(* Logix 5000 project; controller CIP_14485201 vendor 1 type 14 code 216 rev 38.11; software revision 38.01; part 3 of 12 *)
(* tags used below, declared in another part *)
   Alarm_Preset_Indx : DINT;   // ALARM TIMER PRESET INDEX POSITION
   Alarm_Timer : TIMER[128];   // ALARM MSGS 1-127 DELAY TIMERS
   Alarm_Timer_Preset : DINT[128];   // ALARM TIMER PRESETS STORAGE
   Bit : BOOL[128];   // BIT
   Integer : DINT[150];   // INTEGER
   Integer_1 : ALIAS FOR Integer[1];   // RECIPE SELECTOR LIST POSITION ALIAS
   Integer_6 : ALIAS FOR Integer[6];   // EDIT RECIPES SELECTOR LIST POSITION ALIAS
   One_Shot : BOOL[128];   // ONE SHOT ARRAY
   OpCode_Pin : DINT[5];   // OPCODE PIN ARRAY
   OpCode_Word : DINT[5,97];   // OPCODE WORD ARRAY
   Panelview : INT[40];   // PANELVIEW CONTROL
   PID2_Output_Memory : REAL;   // SUPPLY FLOW PID OUTPUT MEMORY TO USE FOR BUMPLESS TRANSFER
   Process_to_CIP : Process_to_CIP;   // PROCESS SIGNALS TO CIP
   PV_Copy_Recipes_Destination : DINT;   // COPY RECIPES DESTINATION
   PV_Copy_Recipes_Duration : TIMER;   // COPY RECIPES COPY DURATION
   PV_Copy_Recipes_One_Shot : BOOL;   // COPY RECIPES REQUEST TO COPY ONE SHOT
   PV_Copy_Recipes_Request : BOOL;   // COPY RECIPES REQUEST TO COPY
   PV_Copy_Recipes_Source : DINT;
   PV_Current_Select_Step_Op : DINT;   // PANELVIEW STORES CURRENT OPCODE NUMBER OF STEP BEING EDITED FOR DISPLAY ON OPCODE LIST SCREEN
   PV_Edit_OpCode_List : DINT[24];   // PANELVIEW RECIPE EDIT OPCODE LIST
   PV_Edit_Opcode_Sel_Top_Row : DINT;   // PANELVIEW RECIPE EDIT OPCODE LIST TOP ROW #
   PV_Edit_Opcodes : DINT[300];   // PANELVIEW BUFFER TO EDIT OPCODES
   PV_Edit_Recipe_Name : STRING;   // SELECTED RECIPE TO EDIT
   PV_Edit_Recipe_Top_Row : DINT;   // PANELVIEW RECIPE EDIT TOP ROW #
   PV_Edit_Recipes : DINT[7];   // PANELVIEW RECIPE EDITING
   PV_Edit_Recipes_0 : ALIAS FOR PV_Edit_Recipes[0];   // EDIT RECIPES STEP NUMBER
   PV_Edit_Recipes_0_Prev : DINT;   // EDIT RECIPE STEP NUMBER PREVIOUS POSITION
   PV_Edit_Screen_Opcodes : DINT[25];   // PANELVIEW RECIPE EDIT DISPLAY OPCODES
   PV_Edit_Setpoints : REAL[97];   // PANELVIEW BUFFER TO EDIT SETPOINTS
   PV_Edit_Times : DINT[300];   // PANELVIEW BUFFER TO EDIT STEP TIMES
   PV_Edit_Times_Indexer : DINT;
   PV_Edit_Times_Minutes : DINT[98];
   PV_Edit_Times_Seconds : DINT[98];
   PV_Rename_Recipe_Name : STRING;   // PANELVIEW RENAME RECIPE NAME
   PV_Step_Time : DINT;   // PANELVIEW DISPLAY STEP TIME
   pv_step_time_minutes : DINT;   // PANELVIEW DISPLAY STEP TIME MINUTES
   pv_step_time_seconds : DINT;   // PANELVIEW DISPLAY STEP TIME SECONDS
   Recipe : RECIPE[41];   // RECIPES
   Recipe_Name : STRING[41];   // RECIPE NAME STORAGE
   Recipe_Name_Indx : DINT;   // RECIPE NAME INDEX POSITION
   Recipe_Step_Length : CONTROL;   // CURRENT RECIPE LENGTH
   Sequencer : CONTROL[4];   // SEQUENCER
   Step_Time_Preset : DINT;
   Subsequent_OpCode_Pin : DINT[5];   // OPCODE PIN ARRAY
   TemporaryRecipeSelection : DINT;
   Time_Date : DINT[20];   // SYSTEM TIME/DATE EDIT/STORAGE
   Timer : TIMER[99];   // TIMER
   Timer_Chem1_Pump : TIMER[7];   // CHEM #1 CONTROL TIMERS
   Timer_Chem2_Pump : TIMER[7];   // CHEM #2 CONTROL TIMERS
   User_Security_Name_Display : STRING;

PROGRAM MainProgram   (* main routine _02_SUB *)

ROUTINE _02_SUB   (* ladder *)
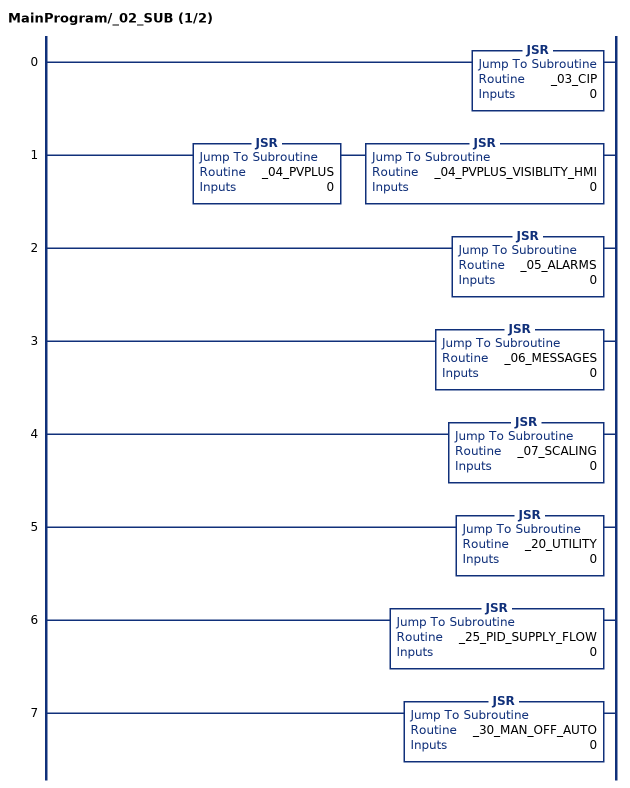
   0: JSR(_03_CIP,0);
   1: JSR(_04_PVPLUS,0)JSR(_04_PVPLUS_VISIBLITY_HMI,0);
   2: JSR(_05_ALARMS,0);
   3: JSR(_06_MESSAGES,0);
   4: JSR(_07_SCALING,0);
   5: JSR(_20_UTILITY,0);
   6: JSR(_25_PID_SUPPLY_FLOW,0);
   7: JSR(_30_MAN_OFF_AUTO,0);
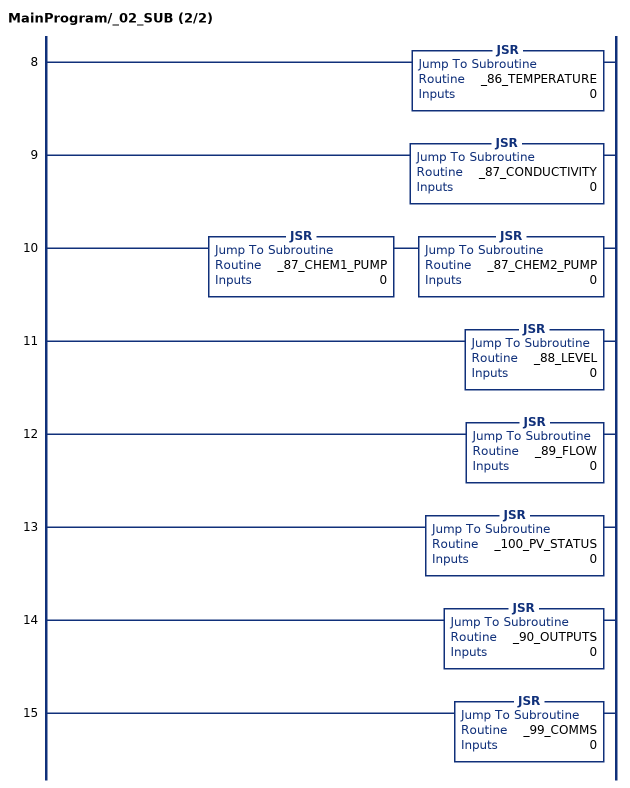
   8: JSR(_86_TEMPERATURE,0);
   9: JSR(_87_CONDUCTIVITY,0);
   10: JSR(_87_CHEM1_PUMP,0)JSR(_87_CHEM2_PUMP,0);
   11: JSR(_88_LEVEL,0);
   12: JSR(_89_FLOW,0);
   13: JSR(_100_PV_STATUS,0);
   14: JSR(_90_OUTPUTS,0);
   15: JSR(_99_COMMS,0);
END_ROUTINE

ROUTINE _03_CIP   (* ladder *)
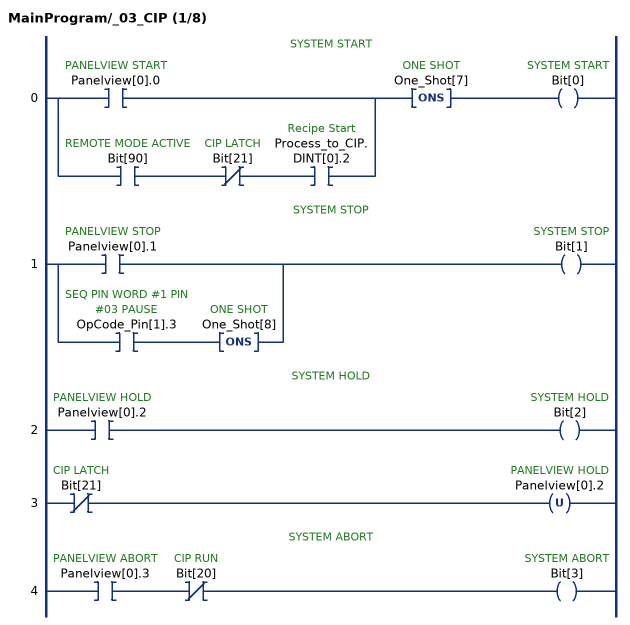
   // SYSTEM START
   0: [XIC(Panelview[0].0) ,XIC(Bit[90]) XIO(Bit[21]) XIC(Process_to_CIP.DINT[0].2) ]ONS(One_Shot[7])OTE(Bit[0]);
   // SYSTEM STOP
   1: [XIC(Panelview[0].1) ,XIC(OpCode_Pin[1].3) ONS(One_Shot[8]) ]OTE(Bit[1]);
   // SYSTEM HOLD
   2: XIC(Panelview[0].2)OTE(Bit[2]);
   3: XIO(Bit[21])OTU(Panelview[0].2);
   // SYSTEM ABORT
   4: XIC(Panelview[0].3)XIO(Bit[20])OTE(Bit[3]);
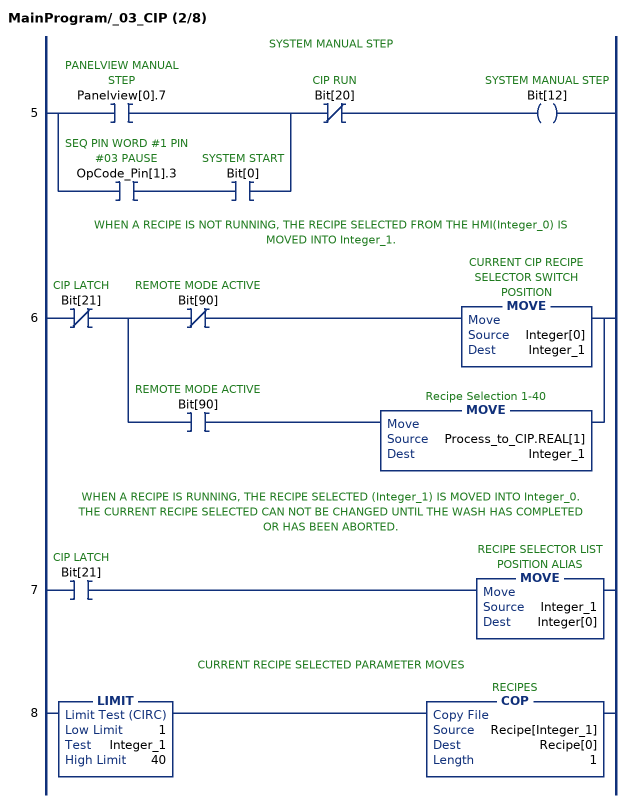
   // SYSTEM MANUAL STEP
   5: [XIC(Panelview[0].7) ,XIC(OpCode_Pin[1].3) XIC(Bit[0]) ]XIO(Bit[20])OTE(Bit[12]);
   // WHEN A RECIPE IS NOT RUNNING, THE RECIPE SELECTED FROM THE HMI(Integer_0) IS MOVED INTO Integer_1.
   6: XIO(Bit[21])[XIO(Bit[90]) MOVE(Integer[0],Integer_1) ,XIC(Bit[90]) MOVE(Process_to_CIP.REAL[1],Integer_1) ];
   // WHEN A RECIPE IS RUNNING, THE RECIPE SELECTED (Integer_1) IS MOVED INTO Integer_0.
   // THE CURRENT RECIPE SELECTED CAN NOT BE CHANGED UNTIL THE WASH HAS COMPLETED OR HAS BEEN ABORTED.
   7: XIC(Bit[21])MOVE(Integer_1,Integer[0]);
   // CURRENT RECIPE SELECTED PARAMETER MOVES
   8: LIMIT(1,Integer_1,40)COP(Recipe[Integer_1],Recipe[0],1);
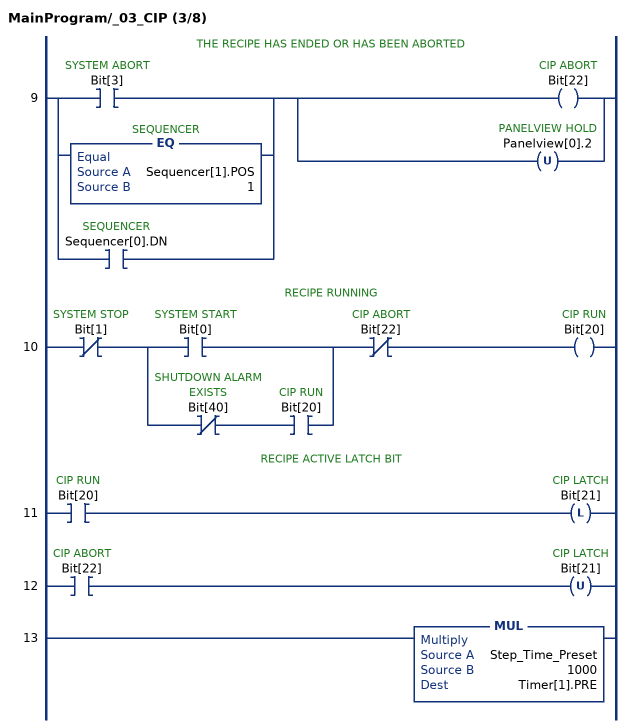
   // THE RECIPE HAS ENDED OR HAS BEEN ABORTED
   9: [XIC(Bit[3]) ,EQ(Sequencer[1].POS,1) ,XIC(Sequencer[0].DN) ][OTE(Bit[22]) ,OTU(Panelview[0].2) ];
   // RECIPE RUNNING
   10: XIO(Bit[1])[XIC(Bit[0]) ,XIO(Bit[40]) XIC(Bit[20]) ]XIO(Bit[22])OTE(Bit[20]);
   // RECIPE ACTIVE LATCH BIT
   11: XIC(Bit[20])OTL(Bit[21]);
   12: XIC(Bit[22])OTU(Bit[21]);
   13: MUL(Step_Time_Preset,1000,Timer[1].PRE);
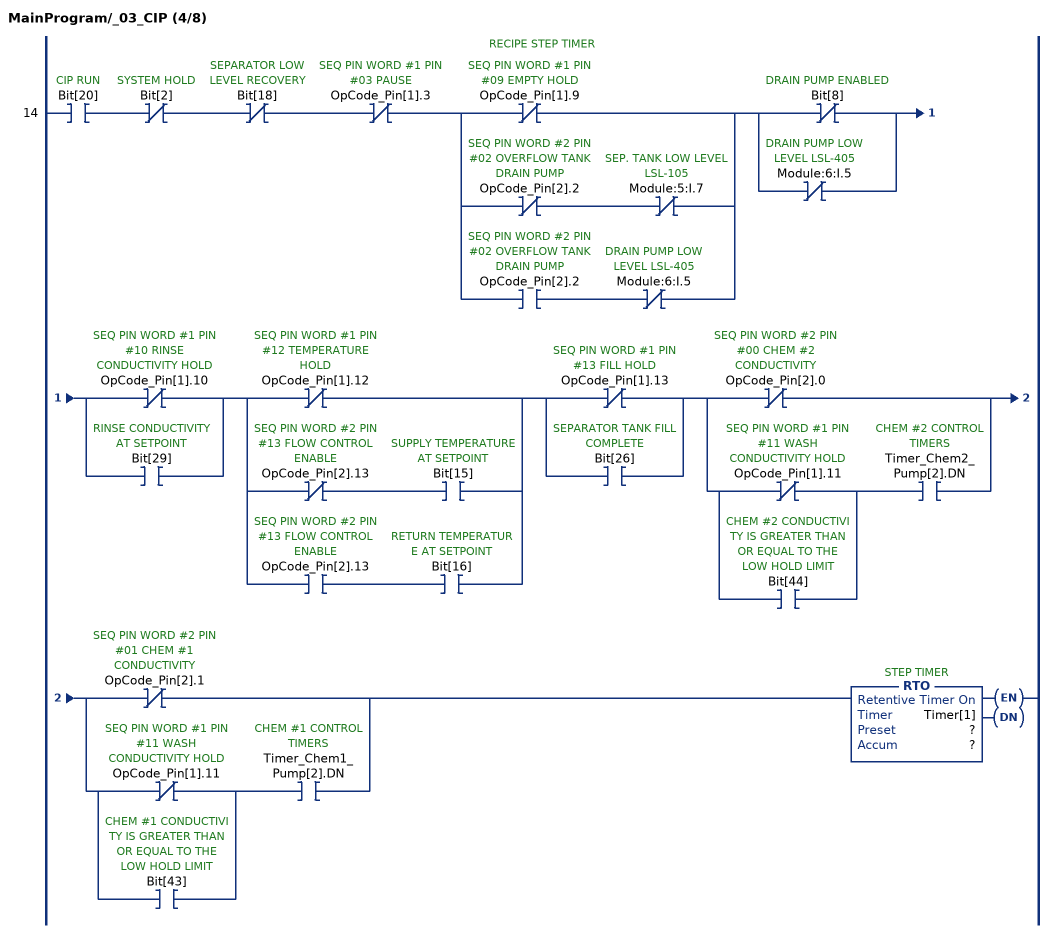
   // RECIPE STEP TIMER
   14: XIC(Bit[20])XIO(Bit[2])XIO(Bit[18])XIO(OpCode_Pin[1].3)[XIO(OpCode_Pin[1].9) ,XIO(OpCode_Pin[2].2) XIO(Module:5:I.7) ,XIC(OpCode_Pin[2].2) XIO(Module:6:I.5) ][XIO(Bit[8]) ,XIO(Module:6:I.5) ][XIO(OpCode_Pin[1].10) ,XIC(Bit[29]) ][XIO(OpCode_Pin[1].12) ,XIO(OpCode_Pin[2].13) XIC(Bit[15]) ,XIC(OpCode_Pin[2].13) XIC(Bit[16]) ][XIO(OpCode_Pin[1].13) ,XIC(Bit[26]) ][XIO(OpCode_Pin[2].0) ,[XIO(OpCode_Pin[1].11) ,XIC(Bit[44]) ] XIC(Timer_Chem2_Pump[2].DN) ][XIO(OpCode_Pin[2].1) ,[XIO(OpCode_Pin[1].11) ,XIC(Bit[43]) ] XIC(Timer_Chem1_Pump[2].DN) ]RTO(Timer[1],?,?);
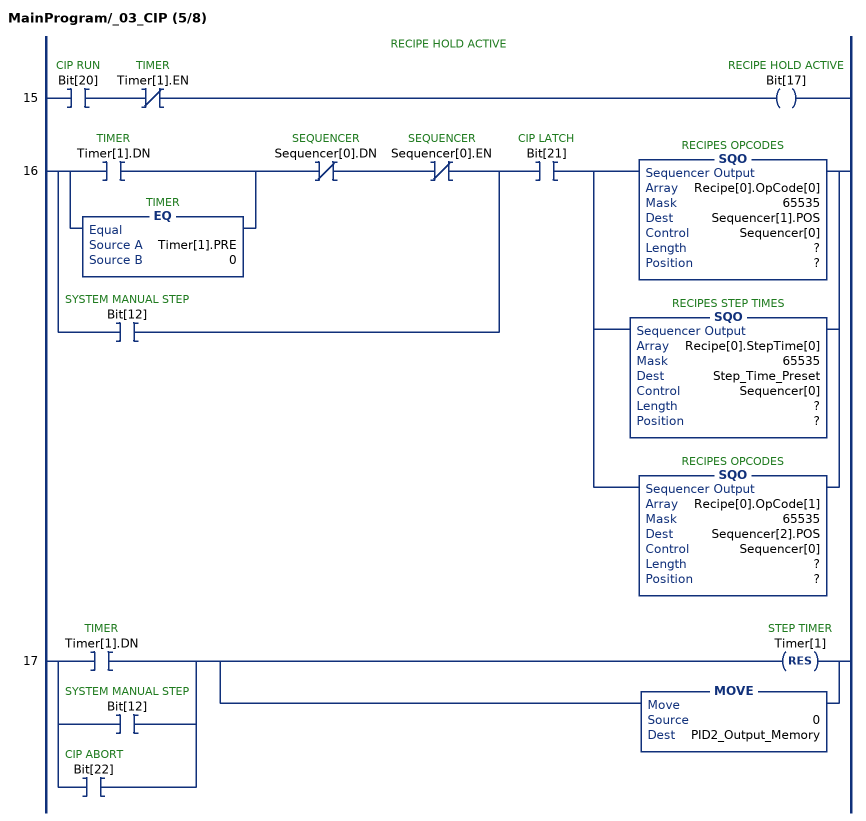
   // RECIPE HOLD ACTIVE
   15: XIC(Bit[20])XIO(Timer[1].EN)OTE(Bit[17]);
   16: [[XIC(Timer[1].DN) ,EQ(Timer[1].PRE,0) ] XIO(Sequencer[0].DN) XIO(Sequencer[0].EN) ,XIC(Bit[12]) ]XIC(Bit[21])[SQO(Recipe[0].OpCode[0],65535,Sequencer[1].POS,Sequencer[0],?,?) ,SQO(Recipe[0].StepTime[0],65535,Step_Time_Preset,Sequencer[0],?,?) ,SQO(Recipe[0].OpCode[1],65535,Sequencer[2].POS,Sequencer[0],?,?) ];
   17: [XIC(Timer[1].DN) ,XIC(Bit[12]) ,XIC(Bit[22]) ][RES(Timer[1]) ,MOVE(0,PID2_Output_Memory) ];
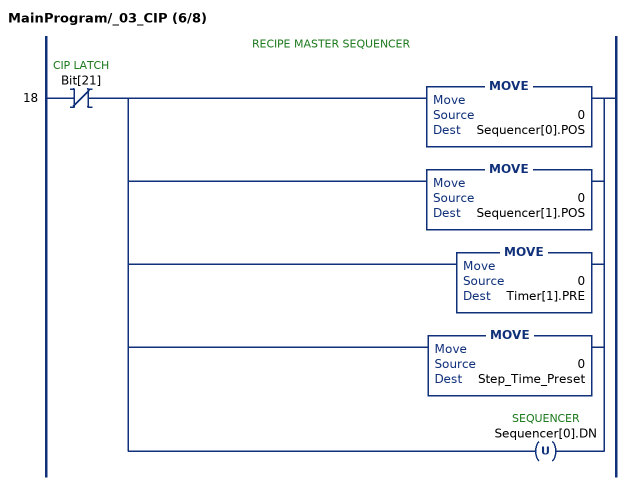
   // RECIPE MASTER SEQUENCER
   18: XIO(Bit[21])[MOVE(0,Sequencer[0].POS) ,MOVE(0,Sequencer[1].POS) ,MOVE(0,Timer[1].PRE) ,MOVE(0,Step_Time_Preset) ,OTU(Sequencer[0].DN) ];
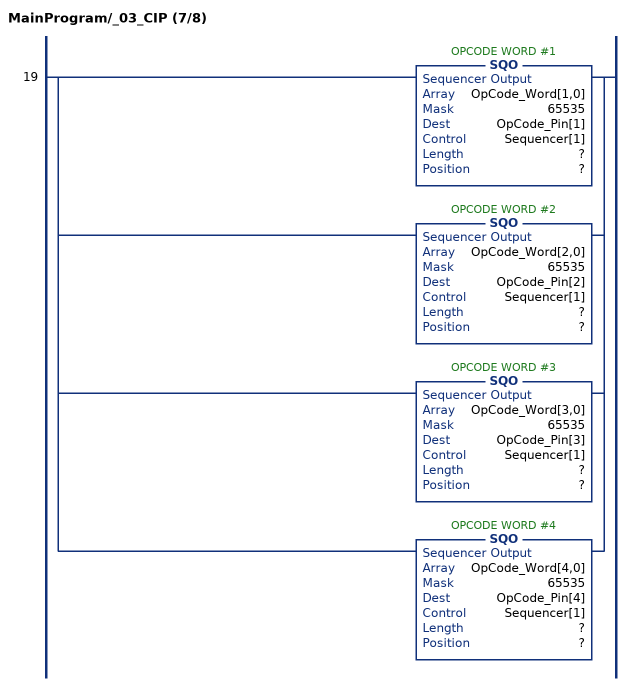
   19: [SQO(OpCode_Word[1,0],65535,OpCode_Pin[1],Sequencer[1],?,?) ,SQO(OpCode_Word[2,0],65535,OpCode_Pin[2],Sequencer[1],?,?) ,SQO(OpCode_Word[3,0],65535,OpCode_Pin[3],Sequencer[1],?,?) ,SQO(OpCode_Word[4,0],65535,OpCode_Pin[4],Sequencer[1],?,?) ];
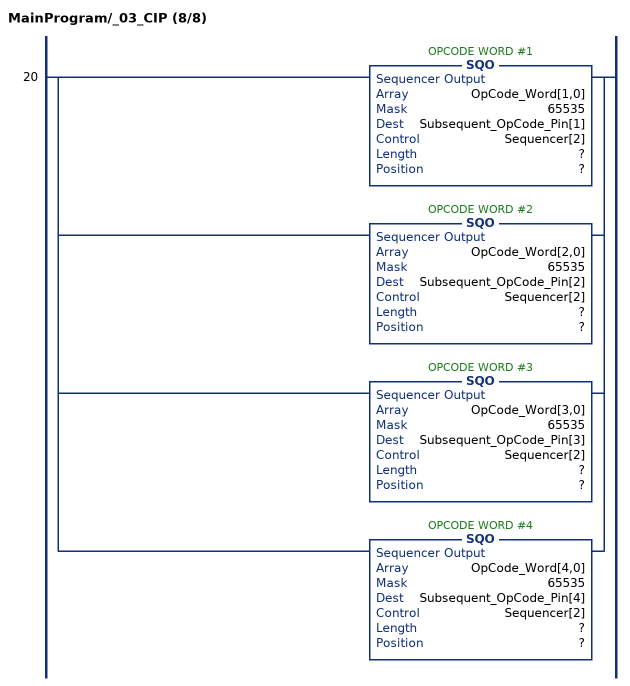
   20: [SQO(OpCode_Word[1,0],65535,Subsequent_OpCode_Pin[1],Sequencer[2],?,?) ,SQO(OpCode_Word[2,0],65535,Subsequent_OpCode_Pin[2],Sequencer[2],?,?) ,SQO(OpCode_Word[3,0],65535,Subsequent_OpCode_Pin[3],Sequencer[2],?,?) ,SQO(OpCode_Word[4,0],65535,Subsequent_OpCode_Pin[4],Sequencer[2],?,?) ];
END_ROUTINE

ROUTINE _04_PVPLUS   (* ladder *)
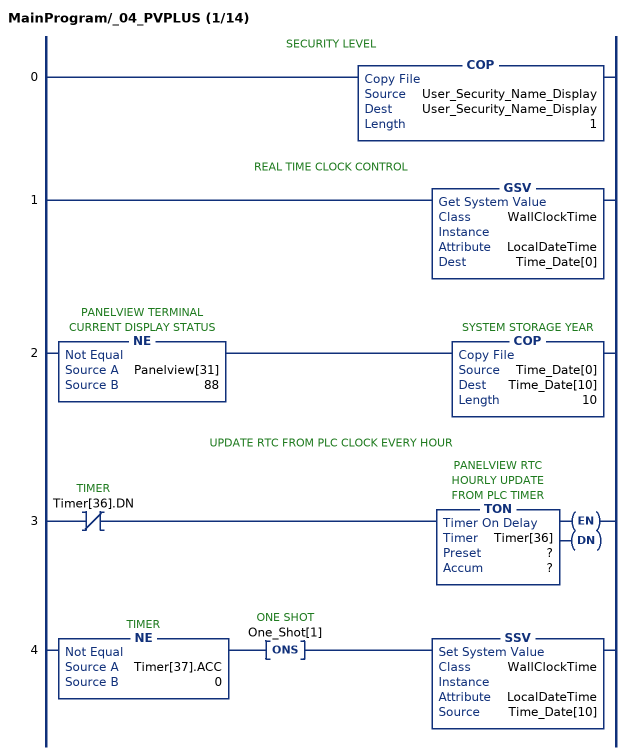
   // SECURITY LEVEL
   0: COP(User_Security_Name_Display,User_Security_Name_Display,1);
   // REAL TIME CLOCK CONTROL
   1: GSV(WallClockTime,,LocalDateTime,Time_Date[0]);
   2: NE(Panelview[31],88)COP(Time_Date[0],Time_Date[10],10);
   // UPDATE RTC FROM PLC CLOCK EVERY HOUR
   3: XIO(Timer[36].DN)TON(Timer[36],?,?);
   4: NE(Timer[37].ACC,0)ONS(One_Shot[1])SSV(WallClockTime,,LocalDateTime,Time_Date[10]);
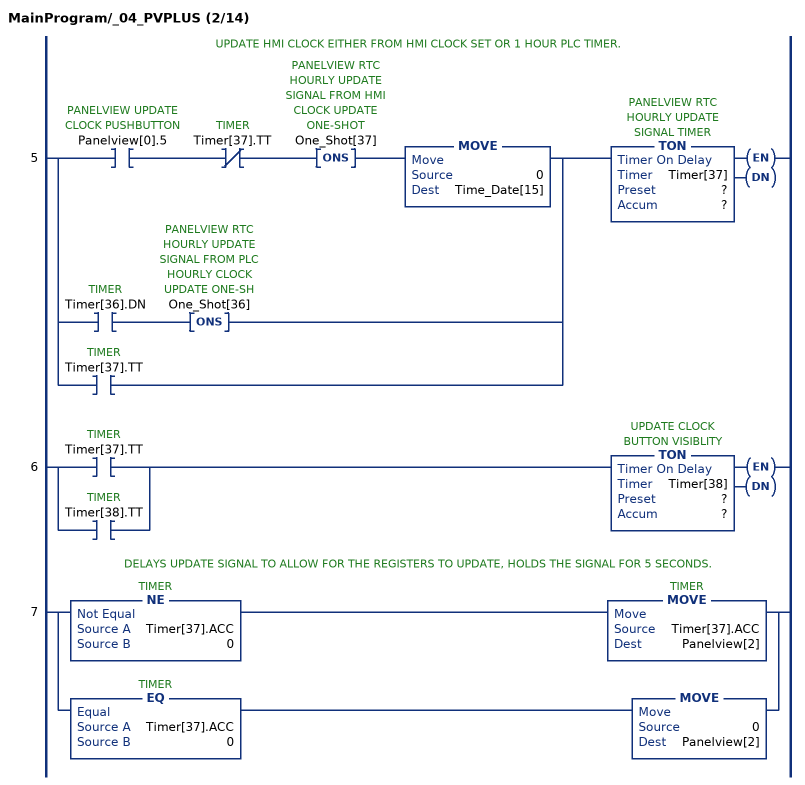
   // UPDATE HMI CLOCK EITHER FROM HMI CLOCK SET OR 1 HOUR PLC TIMER.
   5: [XIC(Panelview[0].5) XIO(Timer[37].TT) ONS(One_Shot[37]) MOVE(0,Time_Date[15]) ,XIC(Timer[36].DN) ONS(One_Shot[36]) ,XIC(Timer[37].TT) ]TON(Timer[37],?,?);
   6: [XIC(Timer[37].TT) ,XIC(Timer[38].TT) ]TON(Timer[38],?,?);
   // DELAYS UPDATE SIGNAL TO ALLOW FOR THE REGISTERS TO UPDATE, HOLDS THE SIGNAL FOR 5 SECONDS.
   7: [NE(Timer[37].ACC,0) MOVE(Timer[37].ACC,Panelview[2]) ,EQ(Timer[37].ACC,0) MOVE(0,Panelview[2]) ];
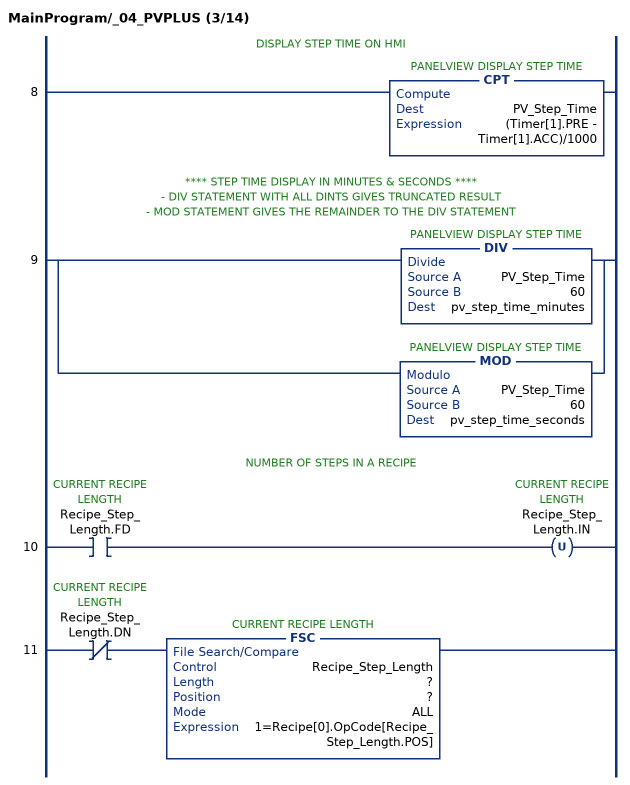
   // DISPLAY STEP TIME ON HMI
   8: CPT(PV_Step_Time,(Timer[1].PRE - Timer[1].ACC)/1000);
   // **** STEP TIME DISPLAY IN MINUTES & SECONDS ****
   // - DIV STATEMENT WITH ALL DINTS GIVES TRUNCATED RESULT
   // - MOD STATEMENT GIVES THE REMAINDER TO THE DIV STATEMENT
   9: [DIV(PV_Step_Time,60,pv_step_time_minutes) ,MOD(PV_Step_Time,60,pv_step_time_seconds) ];
   // NUMBER OF STEPS IN A RECIPE
   10: XIC(Recipe_Step_Length.FD)OTU(Recipe_Step_Length.IN);
   11: XIO(Recipe_Step_Length.DN)FSC(Recipe_Step_Length,?,?,ALL,1=Recipe[0].OpCode[Recipe_Step_Length.POS]);
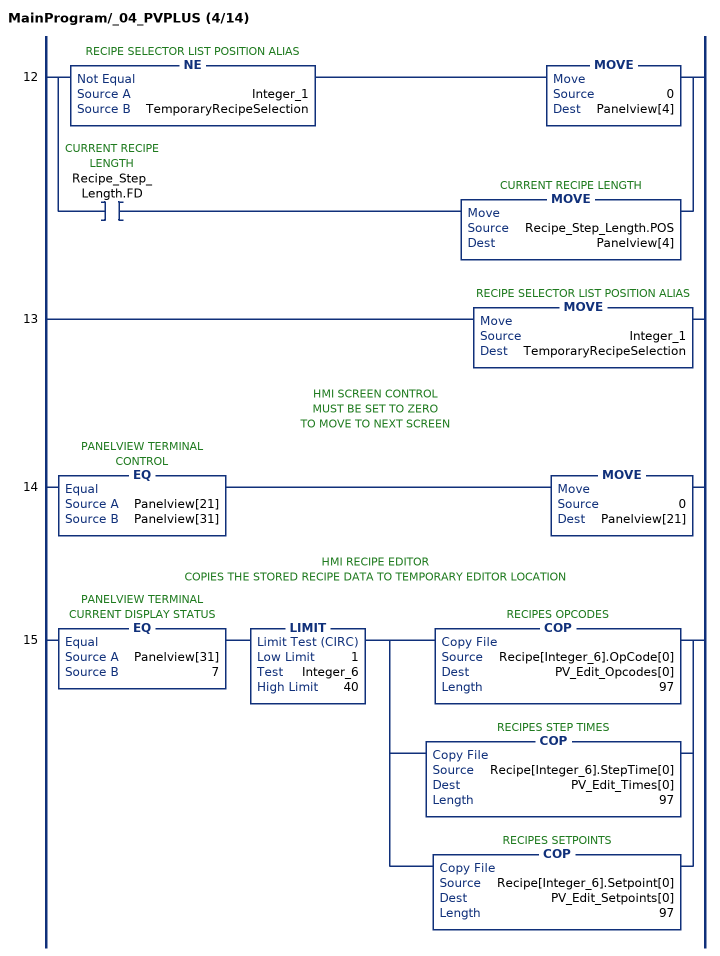
   12: [NE(Integer_1,TemporaryRecipeSelection) MOVE(0,Panelview[4]) ,XIC(Recipe_Step_Length.FD) MOVE(Recipe_Step_Length.POS,Panelview[4]) ];
   13: MOVE(Integer_1,TemporaryRecipeSelection);
   // HMI SCREEN CONTROL
   // MUST BE SET TO ZERO
   // TO MOVE TO NEXT SCREEN
   14: EQ(Panelview[21],Panelview[31])MOVE(0,Panelview[21]);
   // HMI RECIPE EDITOR
   // COPIES THE STORED RECIPE DATA TO TEMPORARY EDITOR LOCATION
   15: EQ(Panelview[31],7)LIMIT(1,Integer_6,40)[COP(Recipe[Integer_6].OpCode[0],PV_Edit_Opcodes[0],97) ,COP(Recipe[Integer_6].StepTime[0],PV_Edit_Times[0],97) ,COP(Recipe[Integer_6].Setpoint[0],PV_Edit_Setpoints[0],97) ];
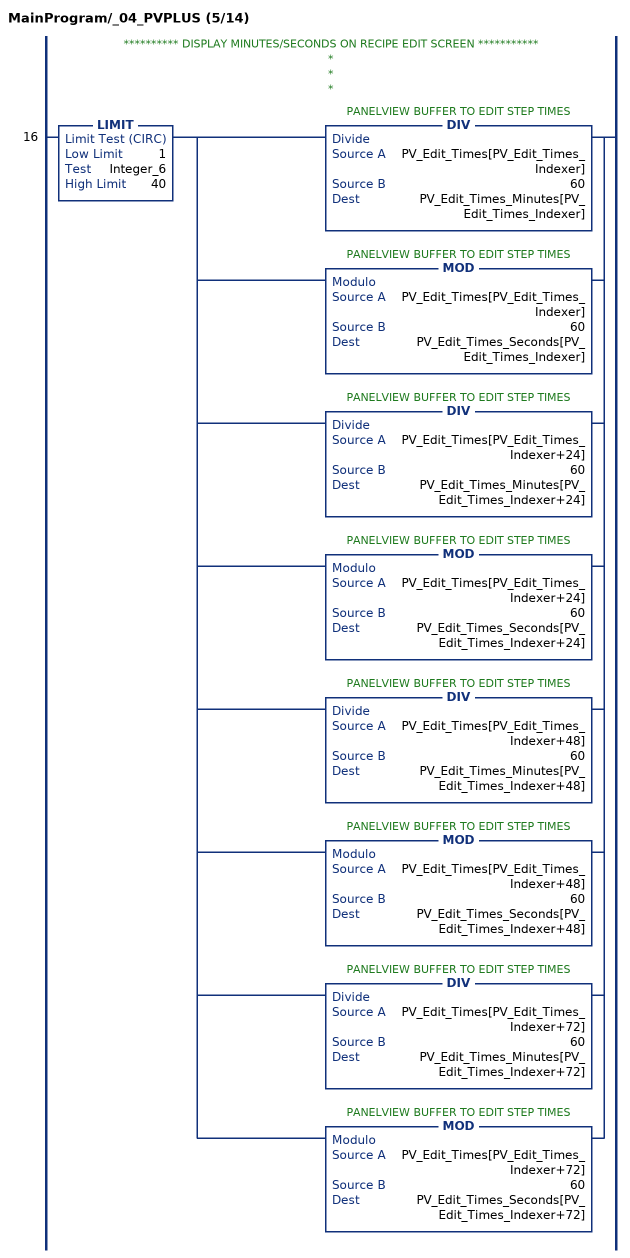
   // ********** DISPLAY MINUTES/SECONDS ON RECIPE EDIT SCREEN ***********
   // *
   // *
   // *
   16: LIMIT(1,Integer_6,40)[DIV(PV_Edit_Times[PV_Edit_Times_Indexer],60,PV_Edit_Times_Minutes[PV_Edit_Times_Indexer]) ,MOD(PV_Edit_Times[PV_Edit_Times_Indexer],60,PV_Edit_Times_Seconds[PV_Edit_Times_Indexer]) ,DIV(PV_Edit_Times[PV_Edit_Times_Indexer+24],60,PV_Edit_Times_Minutes[PV_Edit_Times_Indexer+24]) ,MOD(PV_Edit_Times[PV_Edit_Times_Indexer+24],60,PV_Edit_Times_Seconds[PV_Edit_Times_Indexer+24]) ,DIV(PV_Edit_Times[PV_Edit_Times_Indexer+48],60,PV_Edit_Times_Minutes[PV_Edit_Times_Indexer+48]) ,MOD(PV_Edit_Times[PV_Edit_Times_Indexer+48],60,PV_Edit_Times_Seconds[PV_Edit_Times_Indexer+48]) ,DIV(PV_Edit_Times[PV_Edit_Times_Indexer+72],60,PV_Edit_Times_Minutes[PV_Edit_Times_Indexer+72]) ,MOD(PV_Edit_Times[PV_Edit_Times_Indexer+72],60,PV_Edit_Times_Seconds[PV_Edit_Times_Indexer+72]) ];
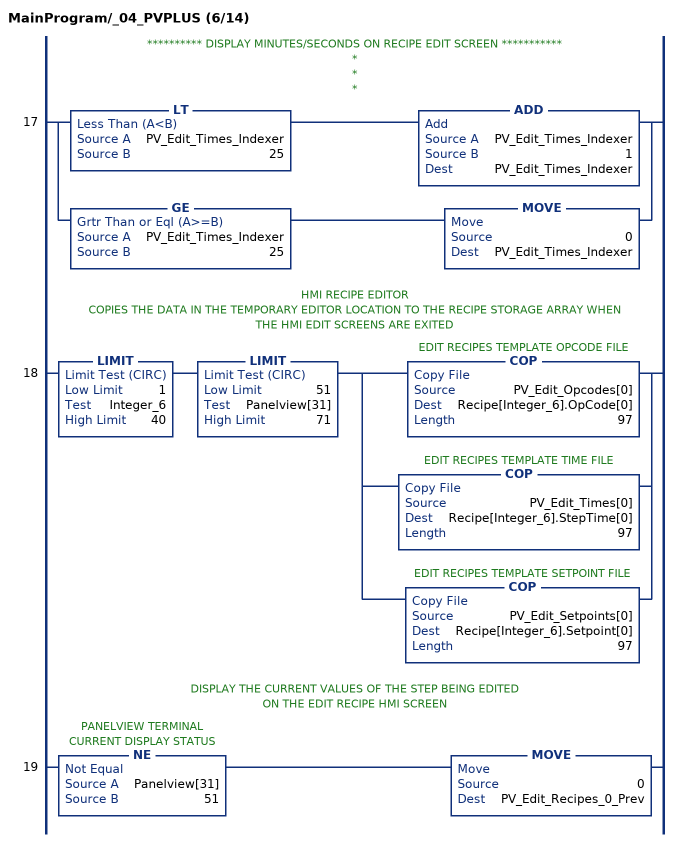
   // ********** DISPLAY MINUTES/SECONDS ON RECIPE EDIT SCREEN ***********
   // *
   // *
   // *
   17: [LT(PV_Edit_Times_Indexer,25) ADD(PV_Edit_Times_Indexer,1,PV_Edit_Times_Indexer) ,GE(PV_Edit_Times_Indexer,25) MOVE(0,PV_Edit_Times_Indexer) ];
   // HMI RECIPE EDITOR
   // COPIES THE DATA IN THE TEMPORARY EDITOR LOCATION TO THE RECIPE STORAGE ARRAY WHEN THE HMI EDIT SCREENS ARE EXITED
   18: LIMIT(1,Integer_6,40)LIMIT(51,Panelview[31],71)[COP(PV_Edit_Opcodes[0],Recipe[Integer_6].OpCode[0],97) ,COP(PV_Edit_Times[0],Recipe[Integer_6].StepTime[0],97) ,COP(PV_Edit_Setpoints[0],Recipe[Integer_6].Setpoint[0],97) ];
   // DISPLAY THE CURRENT VALUES OF THE STEP BEING EDITED
   // ON THE EDIT RECIPE HMI SCREEN
   19: NE(Panelview[31],51)MOVE(0,PV_Edit_Recipes_0_Prev);
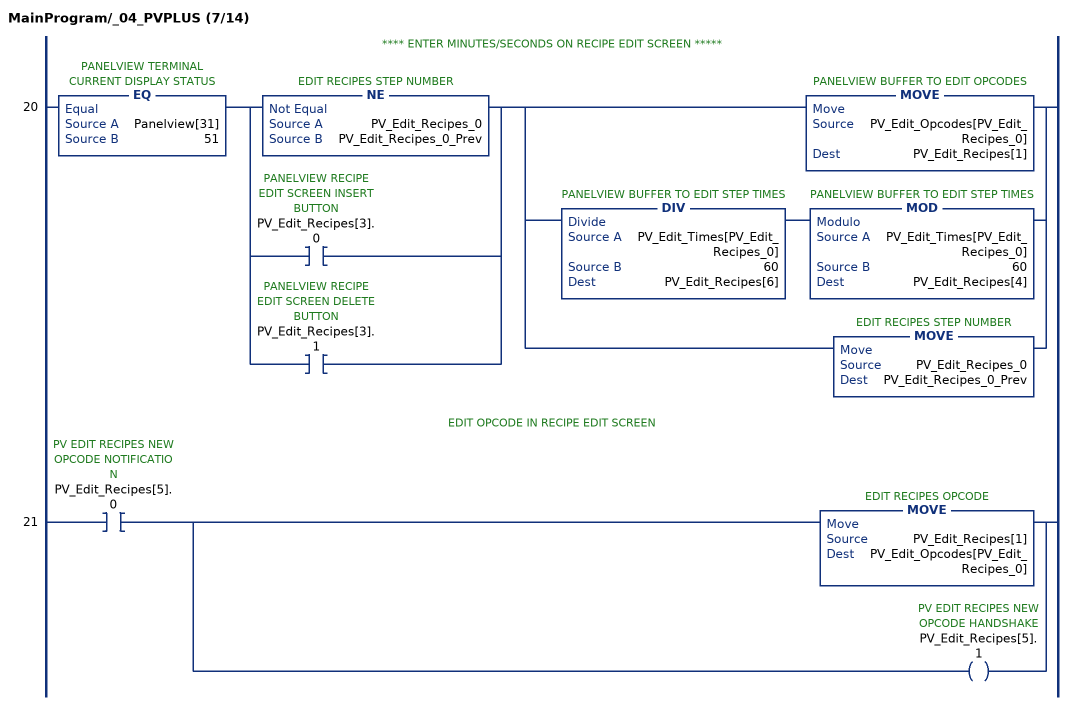
   // **** ENTER MINUTES/SECONDS ON RECIPE EDIT SCREEN *****
   20: EQ(Panelview[31],51)[NE(PV_Edit_Recipes_0,PV_Edit_Recipes_0_Prev) ,XIC(PV_Edit_Recipes[3].0) ,XIC(PV_Edit_Recipes[3].1) ][MOVE(PV_Edit_Opcodes[PV_Edit_Recipes_0],PV_Edit_Recipes[1]) ,DIV(PV_Edit_Times[PV_Edit_Recipes_0],60,PV_Edit_Recipes[6]) MOD(PV_Edit_Times[PV_Edit_Recipes_0],60,PV_Edit_Recipes[4]) ,MOVE(PV_Edit_Recipes_0,PV_Edit_Recipes_0_Prev) ];
   // EDIT OPCODE IN RECIPE EDIT SCREEN
   21: XIC(PV_Edit_Recipes[5].0)[MOVE(PV_Edit_Recipes[1],PV_Edit_Opcodes[PV_Edit_Recipes_0]) ,OTE(PV_Edit_Recipes[5].1) ];
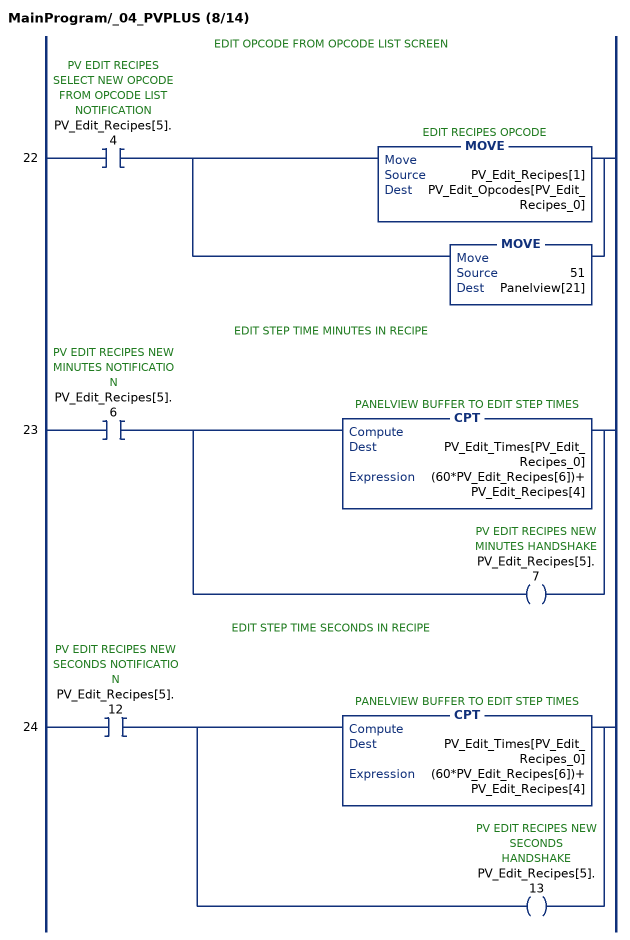
   // EDIT OPCODE FROM OPCODE LIST SCREEN
   22: XIC(PV_Edit_Recipes[5].4)[MOVE(PV_Edit_Recipes[1],PV_Edit_Opcodes[PV_Edit_Recipes_0]) ,MOVE(51,Panelview[21]) ];
   // EDIT STEP TIME MINUTES IN RECIPE
   23: XIC(PV_Edit_Recipes[5].6)[CPT(PV_Edit_Times[PV_Edit_Recipes_0],(60*PV_Edit_Recipes[6])+ PV_Edit_Recipes[4]) ,OTE(PV_Edit_Recipes[5].7) ];
   // EDIT STEP TIME SECONDS IN RECIPE
   24: XIC(PV_Edit_Recipes[5].12)[CPT(PV_Edit_Times[PV_Edit_Recipes_0],(60*PV_Edit_Recipes[6])+ PV_Edit_Recipes[4]) ,OTE(PV_Edit_Recipes[5].13) ];
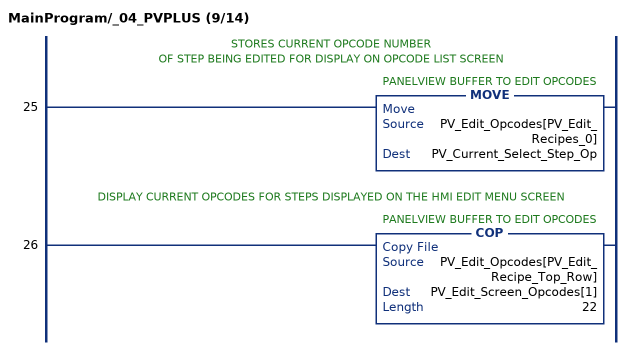
   // STORES CURRENT OPCODE NUMBER
   // OF STEP BEING EDITED FOR DISPLAY ON OPCODE LIST SCREEN
   25: MOVE(PV_Edit_Opcodes[PV_Edit_Recipes_0],PV_Current_Select_Step_Op);
   // DISPLAY CURRENT OPCODES FOR STEPS DISPLAYED ON THE HMI EDIT MENU SCREEN
   26: COP(PV_Edit_Opcodes[PV_Edit_Recipe_Top_Row],PV_Edit_Screen_Opcodes[1],22);
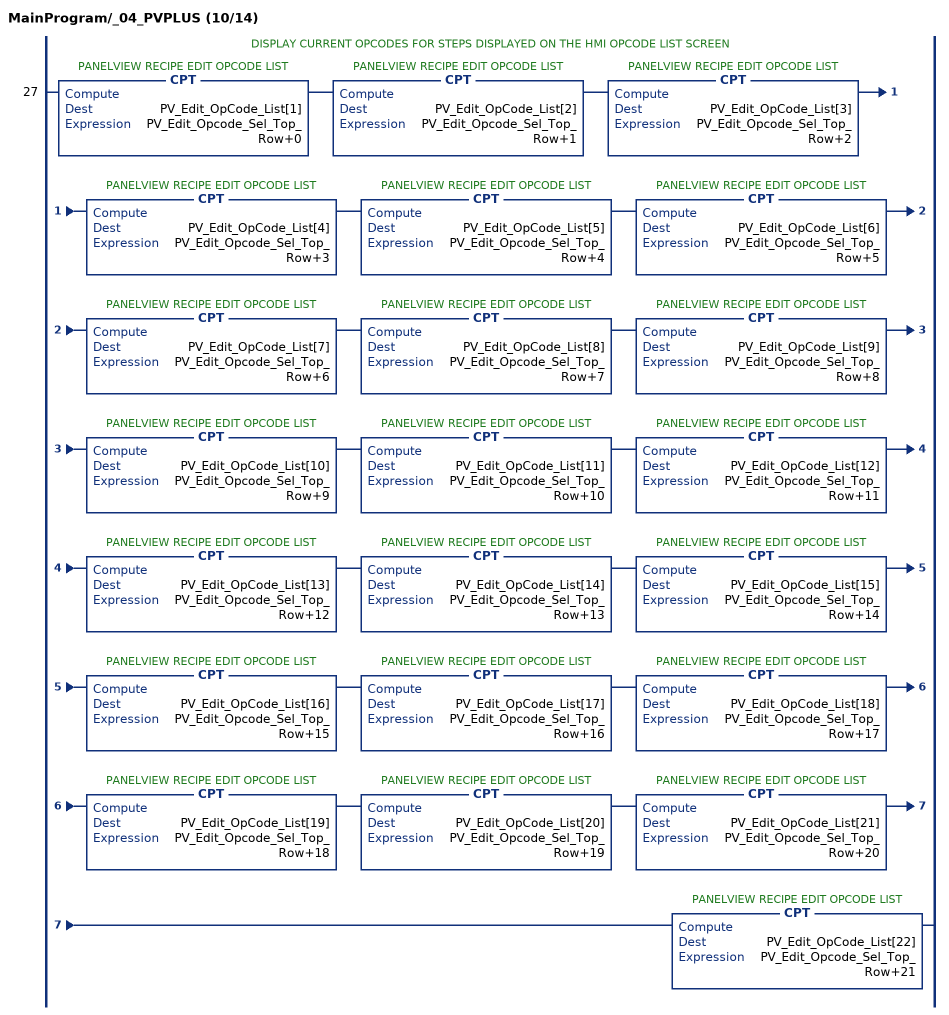
   // DISPLAY CURRENT OPCODES FOR STEPS DISPLAYED ON THE HMI OPCODE LIST SCREEN
   27: CPT(PV_Edit_OpCode_List[1],PV_Edit_Opcode_Sel_Top_Row+0)CPT(PV_Edit_OpCode_List[2],PV_Edit_Opcode_Sel_Top_Row+1)CPT(PV_Edit_OpCode_List[3],PV_Edit_Opcode_Sel_Top_Row+2)CPT(PV_Edit_OpCode_List[4],PV_Edit_Opcode_Sel_Top_Row+3)CPT(PV_Edit_OpCode_List[5],PV_Edit_Opcode_Sel_Top_Row+4)CPT(PV_Edit_OpCode_List[6],PV_Edit_Opcode_Sel_Top_Row+5)CPT(PV_Edit_OpCode_List[7],PV_Edit_Opcode_Sel_Top_Row+6)CPT(PV_Edit_OpCode_List[8],PV_Edit_Opcode_Sel_Top_Row+7)CPT(PV_Edit_OpCode_List[9],PV_Edit_Opcode_Sel_Top_Row+8)CPT(PV_Edit_OpCode_List[10],PV_Edit_Opcode_Sel_Top_Row+9)CPT(PV_Edit_OpCode_List[11],PV_Edit_Opcode_Sel_Top_Row+10)CPT(PV_Edit_OpCode_List[12],PV_Edit_Opcode_Sel_Top_Row+11)CPT(PV_Edit_OpCode_List[13],PV_Edit_Opcode_Sel_Top_Row+12)CPT(PV_Edit_OpCode_List[14],PV_Edit_Opcode_Sel_Top_Row+13)CPT(PV_Edit_OpCode_List[15],PV_Edit_Opcode_Sel_Top_Row+14)CPT(PV_Edit_OpCode_List[16],PV_Edit_Opcode_Sel_Top_Row+15)CPT(PV_Edit_OpCode_List[17],PV_Edit_Opcode_Sel_Top_Row+16)CPT(PV_Edit_OpCode_List[18],PV_Edit_Opcode_Sel_Top_Row+17)CPT(PV_Edit_OpCode_List[19],PV_Edit_Opcode_Sel_Top_Row+18)CPT(PV_Edit_OpCode_List[20],PV_Edit_Opcode_Sel_Top_Row+19)CPT(PV_Edit_OpCode_List[21],PV_Edit_Opcode_Sel_Top_Row+20)CPT(PV_Edit_OpCode_List[22],PV_Edit_Opcode_Sel_Top_Row+21);
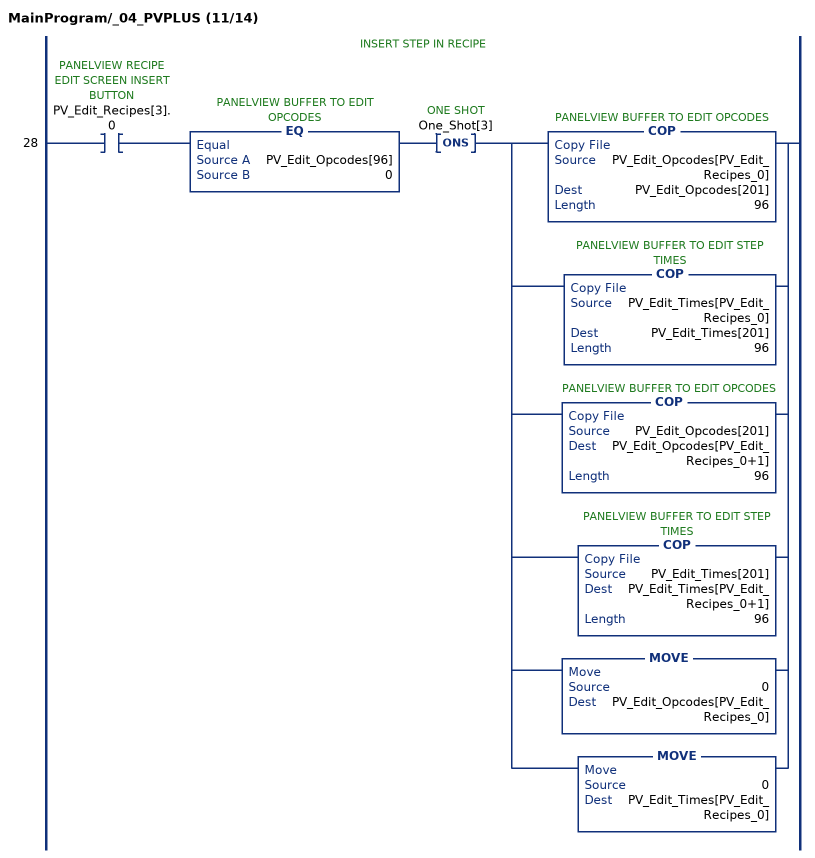
   // INSERT STEP IN RECIPE
   28: XIC(PV_Edit_Recipes[3].0)EQ(PV_Edit_Opcodes[96],0)ONS(One_Shot[3])[COP(PV_Edit_Opcodes[PV_Edit_Recipes_0],PV_Edit_Opcodes[201],96) ,COP(PV_Edit_Times[PV_Edit_Recipes_0],PV_Edit_Times[201],96) ,COP(PV_Edit_Opcodes[201],PV_Edit_Opcodes[PV_Edit_Recipes_0+1],96) ,COP(PV_Edit_Times[201],PV_Edit_Times[PV_Edit_Recipes_0+1],96) ,MOVE(0,PV_Edit_Opcodes[PV_Edit_Recipes_0]) ,MOVE(0,PV_Edit_Times[PV_Edit_Recipes_0]) ];
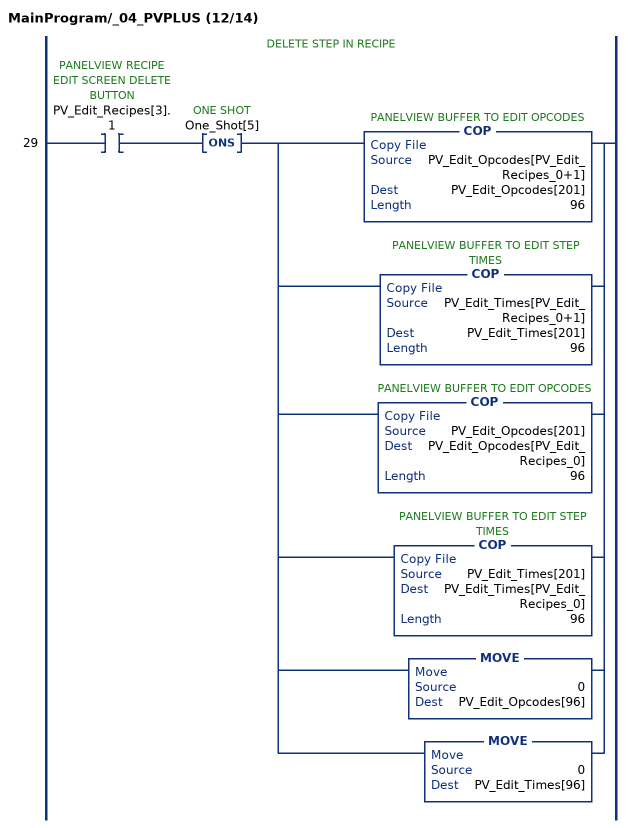
   // DELETE STEP IN RECIPE
   29: XIC(PV_Edit_Recipes[3].1)ONS(One_Shot[5])[COP(PV_Edit_Opcodes[PV_Edit_Recipes_0+1],PV_Edit_Opcodes[201],96) ,COP(PV_Edit_Times[PV_Edit_Recipes_0+1],PV_Edit_Times[201],96) ,COP(PV_Edit_Opcodes[201],PV_Edit_Opcodes[PV_Edit_Recipes_0],96) ,COP(PV_Edit_Times[201],PV_Edit_Times[PV_Edit_Recipes_0],96) ,MOVE(0,PV_Edit_Opcodes[96]) ,MOVE(0,PV_Edit_Times[96]) ];
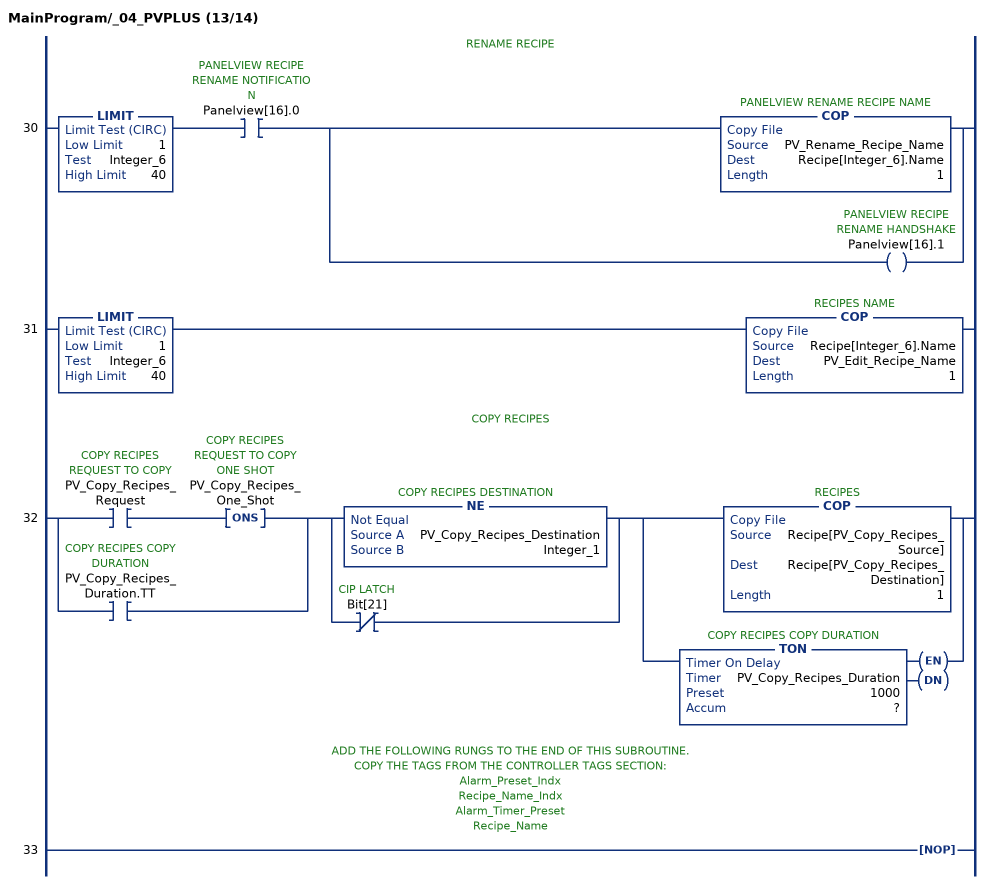
   // RENAME RECIPE
   30: LIMIT(1,Integer_6,40)XIC(Panelview[16].0)[COP(PV_Rename_Recipe_Name,Recipe[Integer_6].Name,1) ,OTE(Panelview[16].1) ];
   31: LIMIT(1,Integer_6,40)COP(Recipe[Integer_6].Name,PV_Edit_Recipe_Name,1);
   // COPY RECIPES
   32: [XIC(PV_Copy_Recipes_Request) ONS(PV_Copy_Recipes_One_Shot) ,XIC(PV_Copy_Recipes_Duration.TT) ][NE(PV_Copy_Recipes_Destination,Integer_1) ,XIO(Bit[21]) ][COP(Recipe[PV_Copy_Recipes_Source],Recipe[PV_Copy_Recipes_Destination],1) ,TON(PV_Copy_Recipes_Duration,?,?) ];
   // ADD THE FOLLOWING RUNGS TO THE END OF THIS SUBROUTINE.
   // COPY THE TAGS FROM THE CONTROLLER TAGS SECTION:
   // Alarm_Preset_Indx
   // Recipe_Name_Indx
   // Alarm_Timer_Preset
   // Recipe_Name
   33: NOP();
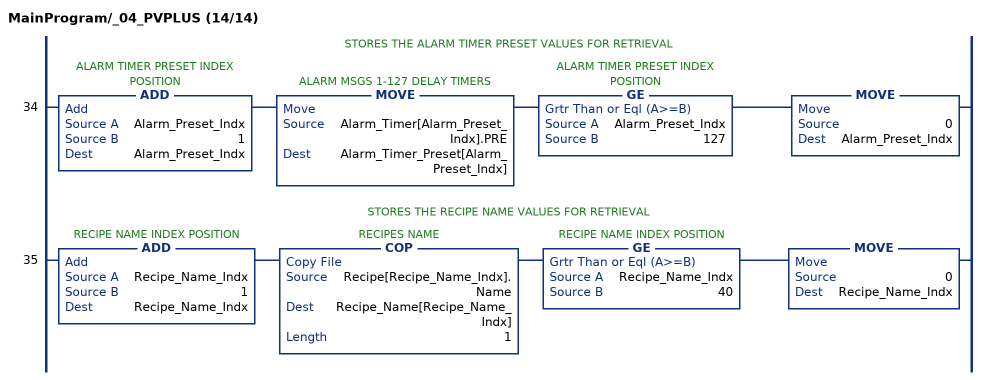
   // STORES THE ALARM TIMER PRESET VALUES FOR RETRIEVAL
   34: ADD(Alarm_Preset_Indx,1,Alarm_Preset_Indx)MOVE(Alarm_Timer[Alarm_Preset_Indx].PRE,Alarm_Timer_Preset[Alarm_Preset_Indx])GE(Alarm_Preset_Indx,127)MOVE(0,Alarm_Preset_Indx);
   // STORES THE RECIPE NAME VALUES FOR RETRIEVAL
   35: ADD(Recipe_Name_Indx,1,Recipe_Name_Indx)COP(Recipe[Recipe_Name_Indx].Name,Recipe_Name[Recipe_Name_Indx],1)GE(Recipe_Name_Indx,40)MOVE(0,Recipe_Name_Indx);
END_ROUTINE
